Fanuc KAREL source: ko00089.KL

-- PROVISIONAL review KL for V1013-1; original PC SHA256 b8b0eb8301b982d7f53153a00523329a5bca2856b9a9b7fc0f275666282d7ddc
-- Incomplete behavior may be omitted. Consult companion uncertainty JSON. Do not deploy.
PROGRAM KO00089
%NOLOCKGROUP
BEGIN
  -- UNRESOLVED_PC offsets 5-12; opcodes 9D,23
  -- UNRESOLVED_PC offsets 17-69; opcodes 27,27,49,7E,AD,27,49,7E,AD,22,31,7E,4A
  -- UNRESOLVED_PC offsets 74-78; opcodes 7F
END KO00089
